(* PLC project probe.project, CODESYS CODESYS V3.5 SP17 Patch 3 *)
(* stored: creationDateTime 2026-10-20T03:54:26.7324602, modificationDateTime 1601-01-01T03:00:00 *)

TYPE ST_ProbeVal : STRUCT
  eMode : E_ProbeMode;
  rValue : REAL := 1.5;
END_STRUCT;
END_TYPE
